// TIA Portal V19 export
DATA_BLOCK "SAFETY"   // DB32
{ S7_Optimized_Access := 'TRUE' }
// stored: MemoryReserve 100
   VAR
      REER_INPUT : "ST_REER_INPUT";
      SAF : "ST_SAF";
      AUTO { S7_SetPoint := 'True'} : Bool;
      MANUAL : Bool;
   END_VAR
BEGIN
END_DATA_BLOCK
